SUBAPPLICATION OptionalGroup_001a (* Optionsgruppe 1a: wie OptionalGroup_001b (Eingang/Ausgang per QI freigeschaltet), reicht die Aktivierung zusaetzlich ueber den Plug PLUG1 an eine nachgeschaltete Gruppe weiter - fuer sequenzielle Aktivierung mehrerer Gruppen (erst 1a, dann 1b). *)
  (* Standard: 61499-2; Description: Copyright (c) 2026 Meisterschulen am Ostbahnhof This program and the accompanying materials are made available under the terms of the Eclipse Public License 2.0 which is available at https://www.eclipse.org/legal/epl-2.0/ SPDX-License-Identifier: EPL-2.0 *)
  (* Version 1.0, 2026-10-13, Franz Höpfinger, Meisterschulen am Ostbahnhof, Daisy-Chain-Glied fuer sequenzielle Options-Aktivierung: PLUG1 (Option::AOption) wird erst ausgeloest, wenn DigitalOutput_Q1 selbst initialisiert ist, und dessen INIT_CNF wird an den eigenen Socket OPTION zurueckgemeldet - der aufrufende DEMUX sieht die Gruppe also erst als fertig, wenn die GESAMTE Kette (inkl. nachgeschalteter Gruppen an PLUG1) bestaetigt hat. *)
  PACKAGE MyLib_AX_Option::sys;
  IMPORT logiBUS::io::DI::logiBUS_DI::Input_I1;
  IMPORT logiBUS::io::DQ::logiBUS_DO::Output_Q1;
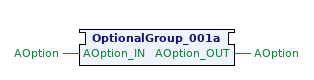
  SOCKETS
    AOption_IN : Option::AOption;
  END_SOCKETS
  PLUGS
    AOption_OUT : Option::AOption;
  END_PLUGS
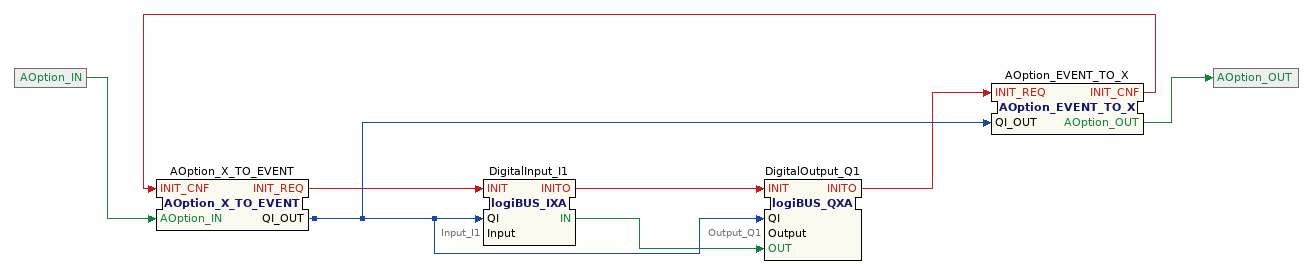
  FBS
    DigitalInput_I1 : logiBUS::io::DI::logiBUS_IXA(Input := Input_I1);
    DigitalOutput_Q1 : logiBUS::io::DQ::logiBUS_QXA(Output := Output_Q1);
    AOption_X_TO_EVENT : Option::conversion::AOption_X_TO_EVENT;
    AOption_EVENT_TO_X : Option::conversion::AOption_EVENT_TO_X;
  END_FBS
  EVENT_CONNECTIONS
    AOption_X_TO_EVENT.INIT_REQ TO DigitalInput_I1.INIT;
    DigitalInput_I1.INITO TO DigitalOutput_Q1.INIT;
    DigitalOutput_Q1.INITO TO AOption_EVENT_TO_X.INIT_REQ;
    AOption_EVENT_TO_X.INIT_CNF TO AOption_X_TO_EVENT.INIT_CNF;
  END_CONNECTIONS
  DATA_CONNECTIONS
    AOption_X_TO_EVENT.QI_OUT TO DigitalInput_I1.QI;
    AOption_X_TO_EVENT.QI_OUT TO DigitalOutput_Q1.QI;
    AOption_X_TO_EVENT.QI_OUT TO AOption_EVENT_TO_X.QI_OUT;
  END_CONNECTIONS
  ADAPTER_CONNECTIONS
    DigitalInput_I1.IN TO DigitalOutput_Q1.OUT;
    AOption_IN TO AOption_X_TO_EVENT.AOption_IN;
    AOption_EVENT_TO_X.AOption_OUT TO AOption_OUT;
  END_CONNECTIONS
END_SUBAPPLICATION
